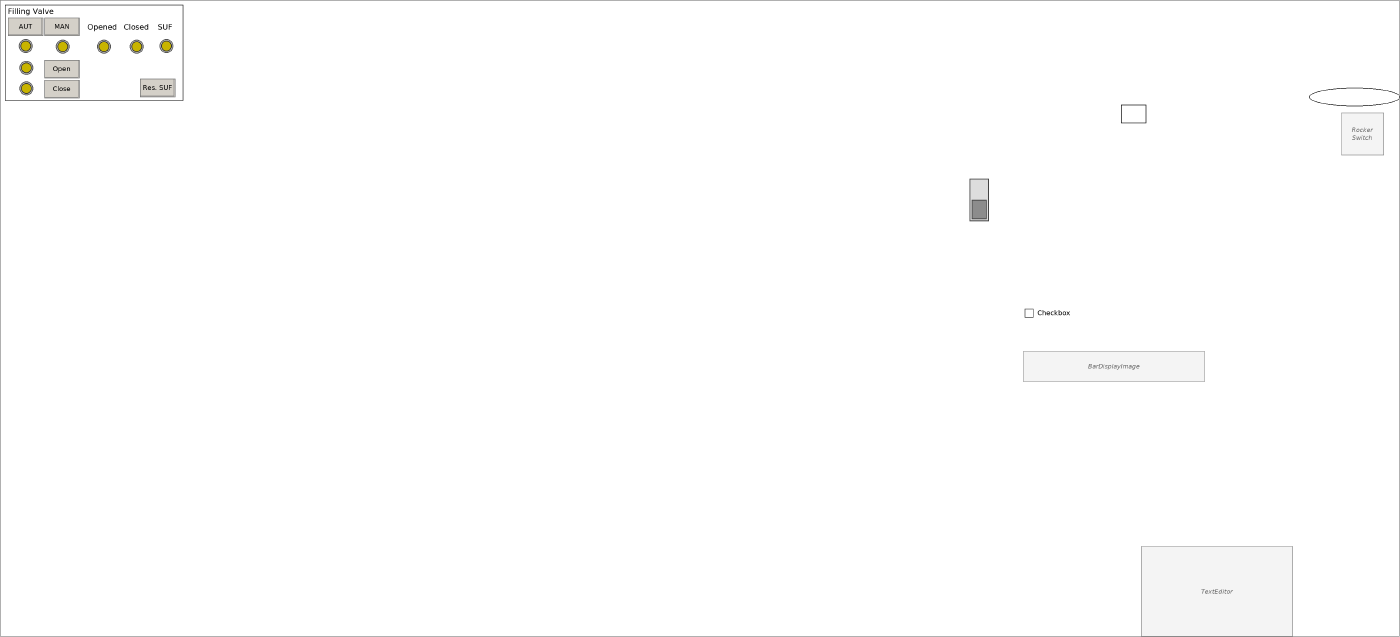
VISUALIZATION Visualization  // 2309x1052
    Rectangle (8,8 294x158)
    Checkbox (1688,502 150x30), "Checkbox"
    BarDisplayImage (1687,580 300x50), style: BarDisplayImage-Gray, scale format: %.1f, scale 0..100
    DipSwitch (1580,295 70x70), behaviour: TOGGLE, style: Switch-DipSwitch-Gray
    RockerSwitch (2212,186 70x70), behaviour: TOGGLE, style: Switch-RockerSwitch-Gray
    TextEditor (1882,902 250x150)
        p4127561890: Courier New
    Ellipse (2159,145 150x30)
    Rectangle (1849,173 41x30)
    Button (13,29 58x30), "AUT"
        OnMouseClick: toggle Global.Tank1.ValveFilling.Cmd.AutCtrl
    Button (73,29 58x30), "MAN"
        OnMouseClick: toggle Global.Tank1.ValveFilling.Cmd.ManCtrl
    Label (10,10 96x18), "Filling Valve"
    Button (73,99 58x30), "Open"
        OnMouseClick: toggle Global.Tank1.ValveFilling.Cmd.OpenMan
    Button (73,132 58x30), "Close"
        OnMouseClick: toggle Global.Tank1.ValveFilling.Cmd.CloseMan
    Lamp1 (29,63 27x26), variable: Global.Tank1.ValveFilling.State.AutCtrl, style: Lamp-Lamp1-Yellow
    Lamp1 (90,64 27x26), variable: Global.Tank1.ValveFilling.State.ManCtrl, style: Lamp-Lamp1-Yellow
    Lamp1 (158,64 27x26), variable: Global.Tank1.ValveFilling.State.Open, style: Lamp-Lamp1-Yellow
    Lamp1 (212,64 27x26), variable: Global.Tank1.ValveFilling.State.Closed, style: Lamp-Lamp1-Yellow
    Lamp1 (261,63 27x26), variable: Global.Tank1.ValveFilling.State.StartupFail, style: Lamp-Lamp1-Yellow
    Button (231,130 58x30), "Res. SUF"
        OnMouseClick: toggle Global.Tank1.ValveFilling.Cmd.ResetSUF
    Label (141,36 53x18), "Opened"
    Label (201,36 53x18), "Closed"
    Label (257,36 33x18), "SUF"
    Lamp1 (30,99 27x26), variable: Global.Tank1.ValveFilling.State.OpenOut, style: Lamp-Lamp1-Yellow
    Lamp1 (30,133 27x26), variable: Global.Tank1.ValveFilling.State.CloseOut, style: Lamp-Lamp1-Yellow
END_VISUALIZATION

(* stored: Version 1.1.0.1, ProductVersion 3.1.4024.13
   Visu Visualization: Id {a6343251-0068-49ba-9adb-31cb88a6e465} *)
